// TIA Portal V21 export
DATA_BLOCK "F_DB_Settings"   // DB7, F_DB
{ S7_Optimized_Access := 'TRUE' }
   VAR
      Signals : "UDT_FSignals";   // Sicherheitssignale / Safety signals
      SetupMode : Bool;   // Einrichtbetrieb angewählt / Setup mode selected
      MachineReleased : Bool;   // Maschine vom Sicherheitsprogramm freigegeben / Machine released by the safety program
   END_VAR
BEGIN
END_DATA_BLOCK
